PROGRAM MAIN
VAR
	//Linking variables to IO cards
	Flow_Valve_1 AT %Q* : INT;
	Level_Valve_1 AT %Q* : INT;
	Level_Valve_2 AT %Q* : INT;
	Level_Valve_3 AT %Q* : INT;
	Gas_Valve AT %Q* : INT;
	Mixer_Valve AT %Q* : INT;
	Motor_speed AT %Q* : INT;
	Motor_ON_OFF AT %Q* :BOOL;
	Motor_Direction AT %Q* :BOOL; 
	Start_Button AT %I* :BOOL;
	Stop_Button AT %I* : BOOL; 
	EMERGENCY_STOP AT %I* : BOOL; 
	Level_Transmitter_1 AT %I* :INT; 
	Level_Transmitter_2 AT %I* :INT; 
	Temperature_Transmitter AT %I* :INT;  
	Pressure_Differencial_Transmitter_1 AT %I* : INT;
	Pressure_Differencial_Transmitter_2 AT %I* : INT;
	Pressure_Transmitter_1 AT %I* : INT ; 
	Pressure_Transmitter_2 AT %I* : INT ; 
	Pressure_Transmitter_3 AT %I* : INT ;
	bSimulate : BOOL := FALSE;   // TRUE = kjører lokalt uten I/O. SETT FALSE PÅ EKTE PLC!
	bReset : BOOL;   // Felles reset fra HMI: alarmer, safe state og motor - olavr

	
	//User Input as percentage
	Flow_Valve_1_Percentage: INT :=100;
	Level_Valve_1_Percentage: INT  := 0;
	Level_Valve_2_Percentage: INT := 0;
	Level_Valve_3_Percentage: INT := 0;
	Motor_speed_Percentage: INT := 0;
	Motor_ON : BOOL ;
	ON_OFF : STRING(10) := 'OFF' ; 
	
	//Scaled values
	Level_Transmitter_1_Scaled : REAL;
	Level_Transmitter_2_Scaled : REAL;
	Pressure_Differential_Transmitter_1_Scaled : REAL;
	Pressure_Differential_Transmitter_2_Scaled : REAL;
	
	//PI function block instantiation
	PI_Controller : PI_Function_Block;
	
	//PI controller on/off state
	bControllerActive : BOOL;
	

    Scale_PT1 : FB_Scale;
	Scale_PT2 : FB_Scale;
	Scale_PT3 : FB_Scale;
	Scale_PDT1: FB_Scale;
	Scale_PDT2: FB_Scale;
    Scale_TT1 : FB_Scale;
	Scale_LT1 : FB_Scale;
	Scale_LT2 : FB_Scale;
    
    Pressure_1_Bar_Scaled : REAL;
	Pressure_2_Bar_Scaled : REAL;
	Pressure_3_Bar_Scaled : REAL;
    Temperature_1_Scaled  : REAL;

	

    bAlarmReset    : BOOL;      // Reset-knapp fra HMI

	fbTempAlarm    : FB_Alarm; // FB_Alarm er røykvarsler-modellen, altså tegningen av hvordan den virker.
	fbPressAlarm   : FB_Alarm;   // fbTempAlarm og fbPressAlarm er to faktiske røykvarslere montert i hvert sitt rom.
	

	// Synlighet for varseltrekant i HMI (trip eller nødstopp) - Variabelen er en string siden HMI
	// Kreven tekst
	
	
	fbEmergency_Shutdown : FB_Emergency_Shutdown;
	
	
	
	// FYSISKE KNAPPER
	fbControlPanel : FB_ControlPanel;
	bHmiStart      : BOOL;
	bHmiStop       : BOOL;
	bHmiEStop      : BOOL;
	
END_VAR

bReset := bAlarmReset OR (Start_Button AND fbEmergency_Shutdown.bTrip);

fbControlPanel(
	bStartPB  := Start_Button,
	bStopPB   := Stop_Button OR bSimulate,
	bEStopPB  := EMERGENCY_STOP OR bSimulate,
	bHmiStart := bHmiStart,
	bHmiStop  := bHmiStop OR fbEmergency_Shutdown.bTrip,
	bHmiEStop := bHmiEStop,
	bReset    := bReset);

// skalerer, regulerer og sender ut signaler

Scale_LT1(RawValue := Level_Transmitter_1, 
          PhysMin := 20.0, 
          PhysMax := 20.5, 
          ScaledValue => Level_Transmitter_1_Scaled);

Scale_LT2(RawValue := Level_Transmitter_2, 
          PhysMin := 50.0, 
          PhysMax := 50.5, 
          ScaledValue => Level_Transmitter_2_Scaled);
		  
// Oppgitt i prosent, fordi de reelle verdiene ikke er kjent.
Scale_PDT1(RawValue := Pressure_Differencial_Transmitter_1, 
          PhysMin := 0.0, 
          PhysMax := 100.0, 
          ScaledValue => Pressure_Differential_Transmitter_1_Scaled);
		  
Scale_PDT2(RawValue := Pressure_Differencial_Transmitter_2, 
          PhysMin := 45.0, 
          PhysMax := 45.5, 
          ScaledValue => Pressure_Differential_Transmitter_2_Scaled);

// Skaler PT1 (f.eks. 0 til 6 bar)
Scale_PT1(RawValue := Pressure_Transmitter_1, 
          PhysMin := 0.0, 
          PhysMax := 6.0, 
          ScaledValue => Pressure_1_Bar_Scaled);
		  
Scale_PT2(RawValue := Pressure_Transmitter_2, 
          PhysMin := 0.0, 
          PhysMax := 6.0, 
          ScaledValue => Pressure_2_Bar_Scaled);
		  
Scale_PT3(RawValue := Pressure_Transmitter_3, 
          PhysMin := 0.0, 
          PhysMax := 6.0, 
          ScaledValue => Pressure_3_Bar_Scaled);

// Skaler TT1 (f.eks. -200 til 850 grader)
Scale_TT1(RawValue := Temperature_Transmitter, 
          PhysMin := -200.0, 
          PhysMax := 850.0, 
          ScaledValue => Temperature_1_Scaled);
		  
// PI-Controller
PI_Controller(Actual := Level_Transmitter_2_scaled,
bEnable := bControllerActive);
Level_Valve_2_Percentage := REAL_TO_INT(PI_Controller.Output);


// variable interval for Flow_Valve_1_Percentage  form 0 to 100  
IF Flow_Valve_1_Percentage > 100 THEN
	Flow_Valve_1_Percentage := 100; 
	ELSE IF Flow_Valve_1_Percentage < 0 THEN 
		Flow_Valve_1_Percentage := 0; 
	END_IF
	
END_IF

// variable interval for Level_Valve_1_Percentage  form 0 to 100  
IF Level_Valve_1_Percentage > 100 THEN
	Level_Valve_1_Percentage := 100; 
	ELSE IF Level_Valve_1_Percentage < 0 THEN 
		Level_Valve_1_Percentage := 0; 
	END_IF
	
END_IF

// variable interval for Level_Valve_2_Percentage  form 0 to 100 
IF Level_Valve_2_Percentage > 100 THEN
	Level_Valve_2_Percentage := 100; 
	ELSE IF Level_Valve_2_Percentage < 0 THEN 
		Level_Valve_2_Percentage := 0; 
	END_IF
	
END_IF

// variable interval for Level_Valve_3_Percentage  form 0 to 100 
IF Level_Valve_3_Percentage > 100 THEN
	Level_Valve_3_Percentage := 100; 
	ELSE IF Level_Valve_3_Percentage < 0 THEN 
		Level_Valve_3_Percentage := 0; 
	END_IF
	
END_IF



// variable interval for Motor_speed_Percentage  form 0 to 100 
IF Motor_speed_Percentage > 100 THEN
	Motor_speed_Percentage := 100; 
	ELSE IF Motor_speed_Percentage < 0 THEN 
		Motor_speed_Percentage := 0; 
	END_IF
	
END_IF

// Motor går når prosessen kjører. Nødstopp/trip håndteres i fbEmergency_Shutdown
Motor_ON_OFF := fbControlPanel.bRunning;

// Flow_Valve_1 calibration
Flow_Valve_1 := REAL_TO_INT (262.14*Flow_Valve_1_Percentage +6553 ); 

// Level_Valve_1 calibration
Level_Valve_1 := REAL_TO_INT(262.14*Level_Valve_1_Percentage +6553);

// Level_Valve_2 calibration
Level_Valve_2 := REAL_TO_INT(262.14*Level_Valve_2_Percentage +6553);

// Level_Valve_3 calibration
Level_Valve_3 := REAL_TO_INT(262.14*Level_Valve_3_Percentage +6553);


// Motor_speed calibration
Motor_speed := REAL_TO_INT(262.14*Motor_speed_Percentage +6553);


fbTempAlarm(rValue := Temperature_1_Scaled, rLimit := 80.0, bReset := bReset);
fbPressAlarm(rValue := MAX(Pressure_1_Bar_Scaled, MAX(Pressure_2_Bar_Scaled, Pressure_3_Bar_Scaled)), rLimit := 4.0, bReset := bReset);

// Alarmhåndtering: sender warnings og trips til EventLogger/HMI
Alarm_System();

	
// Safe state
fbEmergency_Shutdown(
	Motor_ON_OFF      := Motor_ON_OFF,
	bControllerActive := bControllerActive,
	Motor_speed       := Motor_speed,
	Gas_Valve         := Gas_Valve,
	Flow_Valve_1      := Flow_Valve_1,
	Level_Valve_1     := Level_Valve_1,
	Level_Valve_2     := Level_Valve_2,
	Level_Valve_3     := Level_Valve_3);

// Motorstatus til HMI (etter safe state, så den viser riktig)
IF Motor_ON_OFF THEN
	Motor_ON := FALSE;
	ON_OFF   := 'MOTOR: ON';
ELSE
	Motor_ON := TRUE;
	ON_OFF   := 'MOTOR: OFF';
END_IF

END_PROGRAM

(* stored: Version 1.1.0.1, ProductVersion 3.1.4026.21
   POU MAIN: Id {75317203-8f43-4932-aa88-c7b05e9ca563}, SpecialFunc None *)
